FUNCTION_BLOCK FB_EmsCmdGate		// EMS command 레코드 앞단: 버전 2 명령을 Delay(ms)만큼 기다렸다가 내보내기
(* 인터페이스 100.Command 버전 2 (2026-11-25): SequenceNumber 없는 16 B 레코드.
   - Delay = 0이면 이번 스캔에 처리한다. Delay > 0이면 보관하고 시간이 되면 핸들러에 넘긴다.
   - 보관 중 같은 장치에 새 명령이 오면 새 명령을 따른다. 1시간을 넘는 Delay는 버린다.
   - 같은 명령을 다시 보내도 처리한다. 재시작하면 보관 중인 명령은 실행하지 않는다. *)
VAR_IN_OUT
	iq_astRec			: ARRAY[*] OF ST_MqttCommand_Rx;	// 수신 배열 (0부터, 칸 = DeviceIndex-1)
END_VAR
VAR_OUTPUT
	q_nDelayedCount		: UDINT;	// Delay 때문에 보관한 수
	q_nReplacedCount	: UDINT;	// 보관 중 새 명령이 와서 버린 보관 명령 수
	q_nBadDelayCount	: UDINT;	// Delay가 너무 커서 버린 수
	q_nPendingCount		: UDINT;	// 지금 보관 중인 명령 수
END_VAR
VAR CONSTANT
	MAX_SLOTS			: DINT := 16;			// 다룰 수 있는 칸 수 (PCS·BMS·UPS 대수보다 커야 함)
	MAX_DELAY_MS		: UDINT := 3600000;		// 1시간
END_VAR
VAR
	_astPend			: ARRAY[0..15] OF ST_MqttCommand_Rx;
	_abPend				: ARRAY[0..15] OF BOOL;
	_atStart			: ARRAY[0..15] OF TIME;
	_tNow				: TIME;
	_i					: DINT;
	_s					: DINT;
END_VAR

_tNow := TIME();
q_nPendingCount := 0;
FOR _i := LOWER_BOUND(iq_astRec, 1) TO UPPER_BOUND(iq_astRec, 1) DO
	_s := _i - LOWER_BOUND(iq_astRec, 1);
	IF _s >= MAX_SLOTS THEN
		EXIT;
	END_IF
	IF iq_astRec[_i].CommandType <> 0 THEN
		IF _abPend[_s] THEN
			_abPend[_s] := FALSE;
			q_nReplacedCount := q_nReplacedCount + 1;
		END_IF
		IF iq_astRec[_i].Delay > MAX_DELAY_MS THEN
			iq_astRec[_i].CommandType := 0;
			q_nBadDelayCount := q_nBadDelayCount + 1;
		ELSIF iq_astRec[_i].Delay > 0 THEN
			_astPend[_s] := iq_astRec[_i];
			_abPend[_s] := TRUE;
			_atStart[_s] := _tNow;
			iq_astRec[_i].CommandType := 0;
			q_nDelayedCount := q_nDelayedCount + 1;
		END_IF
	ELSIF _abPend[_s] AND (_tNow - _atStart[_s]) >= UDINT_TO_TIME(_astPend[_s].Delay) THEN
		iq_astRec[_i] := _astPend[_s];			// 시간이 됨: 이번 스캔에 핸들러가 처리
		iq_astRec[_i].Delay := 0;
		_abPend[_s] := FALSE;
	END_IF
	IF _abPend[_s] THEN
		q_nPendingCount := q_nPendingCount + 1;
	END_IF
END_FOR

END_FUNCTION_BLOCK

(* stored: Version 1.1.0.1, ProductVersion 3.1.4024.12
   POU FB_EmsCmdGate: Id {5f94382c-e185-4e4a-8fb1-a6c5bf5441a8}, SpecialFunc None *)
